FUNCTION_BLOCK FB_ProcessControl

VAR_IN_OUT
	stProcessControl	:	ST_ProcessControl	;
END_VAR
VAR
	bRun			: BOOL	;
	//fbPID	: 	FB_BasicPID	;
	fbPID	: 	PID	;
	hystCIP_SetPoint: FB_Hysteresis_REAL;
	Call_ActDelayTON	: TON	;
	bRunCalled		: BOOL	;//mRun was called since the last body call

	handling_PID_Manual: TON;

END_VAR

//stProcessControl.bManual:=TRUE;



//Deactivate control 1s after mRun stops being called (body may be called several times per cycle)
Call_ActDelayTON(IN:=stProcessControl.bActiveCntr AND NOT bRunCalled , PT:=T#1S , Q=> , ET=> );
bRunCalled:=FALSE;

m_Check();

act_Call_PID();
act_CallHyst();

handling_PID_Manual(PT:=T#0.5S);//, IN:=TRUE
IF handling_PID_Manual.Q THEN;
	stProcessControl.bManual:=TRUE;
ELSE;
	stProcessControl.bManual:=FALSE;
END_IF

ACTION act_Call_PID:
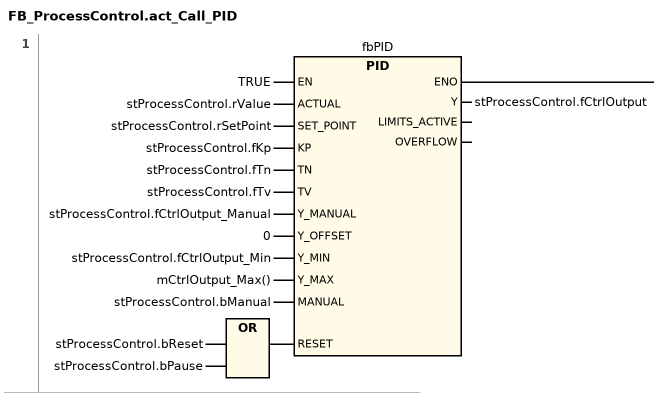
// NETWORK 1
fbPID(
    ACTUAL := stProcessControl.rValue,
    SET_POINT := stProcessControl.rSetPoint,
    KP := stProcessControl.fKp,
    TN := stProcessControl.fTn,
    TV := stProcessControl.fTv,
    Y_MANUAL := stProcessControl.fCtrlOutput_Manual,
    Y_OFFSET := 0,
    Y_MIN := stProcessControl.fCtrlOutput_Min,
    Y_MAX := mCtrlOutput_Max(),
    MANUAL := stProcessControl.bManual,
    RESET := stProcessControl.bReset OR stProcessControl.bPause,
    Y => stProcessControl.fCtrlOutput); // PID
END_ACTION

ACTION act_Call_PID_old:

	
(*
fbPID(
	fSetpointValue:=stProcessControl.rSetPoint , 
	fActualValue:=stProcessControl.rValue , 
	bReset:=stProcessControl.bReset , 
	fCtrlCycleTime:=stProcessControl.fCtrlCycleTime , 
	fKp:=stProcessControl.fKp , 
	fTn:=stProcessControl.fTn , 
	fTv:=stProcessControl.fTv , 
	fTd:=stProcessControl.fTd , 
	fCtrlOutput=>stProcessControl.fCtrlOutput , 
	nErrorStatus=>stProcessControl.nErrorStatus );
*)
END_ACTION

ACTION act_CallHyst:
hystCIP_SetPoint(
	fIn:=stProcessControl.rValue,//g_HMI.stT4_Sens.rTankLevel,
	fHigh:=stProcessControl.fHystHigh,
	fLow:=stProcessControl.fHystLow,
	iDigitsAfterDot:=,
	bOut=>stProcessControl.bHystOut);
END_ACTION

METHOD m_Check : BOOL
VAR_INPUT
END_VAR
IF NOT __ISVALIDREF(stProcessControl) THEN
	RETURN;
END_IF

IF bRun THEN
	stProcessControl.bActiveCntr:=TRUE;
	bRunCalled:=TRUE;
ELSIF NOT bRun AND Call_ActDelayTON.Q THEN
	stProcessControl.bActiveCntr:=FALSE;
END_IF

IF bRun THEN
	stProcessControl.Deviation:=stProcessControl.rSetPoint-stProcessControl.rValue;
	stProcessControl.Control_ON:=FALSE;
	stProcessControl.OverFlow:=FALSE;
	stProcessControl.bDone:=FALSE;
	
	IF stProcessControl.Deviation >= stProcessControl.ToleravceLow THEN;
		//Value too low needs to be increased
		stProcessControl.Control_ON:=TRUE;
		stProcessControl.OverFlow:=FALSE;
		stProcessControl.bDone:=FALSE;
	ELSIF stProcessControl.Deviation <= -stProcessControl.ToleranceHigh THEN;
		//value too high need to be decreased
		stProcessControl.OverFlow:=TRUE;
		stProcessControl.Control_ON:=TRUE;
		stProcessControl.bDone:=FALSE;
		//message
	ELSE;
		// Done, value in tolerace
		stProcessControl.OverFlow:=FALSE;
		stProcessControl.Control_ON:=FALSE;
		stProcessControl.bDone:=TRUE;
	END_IF
	bRun:=FALSE;
END_IF
END_METHOD

METHOD mCtrlOutput_Max : REAL
VAR_INPUT
END_VAR

VAR
	span: LREAL;
END_VAR


span:=ABS(stProcessControl.fCtrlOutput_Max-stProcessControl.fCtrlOutput_Min);
//LimitedPrecentage:=
IF stProcessControl.rValue>stProcessControl.rValue_Min_To_ReleaseControl THEN;
	mCtrlOutput_Max:=stProcessControl.fCtrlOutput_Max;
ELSE;
	mCtrlOutput_Max:=stProcessControl.fCtrlOutput_Min+(span*0.3);
END_IF
END_METHOD

METHOD mManual : BOOL
VAR_INPUT
	value: BOOL;
END_VAR
//PID manual request without starting control (bRun/bActiveCntr untouched)
handling_PID_Manual(IN:=value);
mManual:=stProcessControl.bManual;
END_METHOD

METHOD mPause : BOOL
VAR_INPUT
	value: BOOL;
END_VAR
stProcessControl.bPause:=value;
END_METHOD

METHOD mReset : BOOL
VAR_INPUT
END_VAR
stProcessControl.Control_ON:=FALSE;
stProcessControl.OverFlow:=FALSE;
stProcessControl.bDone:=FALSE;
END_METHOD

METHOD mRun : BOOL
VAR_INPUT
	//Set_Point: REAL;
END_VAR
bRun:=TRUE;
//stProcessControl.rSetPoint:=Set_Point;
m_Check();



mRun:=stProcessControl.bDone;
END_METHOD

METHOD mRun_Hyst : REAL
VAR_INPUT
END_VAR
stProcessControl.bManual:=FALSE;
IF stProcessControl.bHystOut THEN
	mRun_Hyst:=stProcessControl.rHystOutLow;
ELSE
	mRun_Hyst:=stProcessControl.rHystOutHigh;
END_IF
END_METHOD

METHOD mRun_PID : REAL
VAR_INPUT
	Set_Point: REAL;
	controlManual: BOOL;
END_VAR
mRun();//mRun(Set_Point:=Set_Point);
//stProcessControl.bManual:=controlManual;
//stProcessControl.rSetPoint:=Set_Point;
handling_PID_Manual(IN:=controlManual);
mRun_PID:=stProcessControl.fCtrlOutput;
END_METHOD

METHOD mRun_With_SP : BOOL
VAR_INPUT
	Set_Point: REAL;
END_VAR
stProcessControl.rSetPoint:=Set_Point;
bRun:=TRUE;
mRun();
//stProcessControl.rSetPoint:=Set_Point;
mRun_With_SP:=stProcessControl.bDone;
END_METHOD

END_FUNCTION_BLOCK

(* stored: Version 1.1.0.1, ProductVersion 3.1.4026.21
   POU FB_ProcessControl: Id {a1972051-d534-4d79-bd7a-71cd1b516897}, SpecialFunc None
   Action act_Call_PID: Id {839fbd4c-e468-439d-b2e8-fa15b4ee659a}
   Action act_Call_PID_old: Id {e29ea305-112b-4479-9e5c-3d503fcea5b6}
   Action act_CallHyst: Id {7f4572c7-9e9a-4bff-b0e0-f6c19cca19c6}
   Method m_Check: Id {b27ec81e-04ce-483d-958b-1ee4b2519c56}
   Method mCtrlOutput_Max: Id {96e0187b-897b-496a-b800-2f20b878b88c}
   Method mManual: Id {1beeeb9a-e732-4638-8ad0-65b51ae96f3a}
   Method mPause: Id {be53090d-a73d-45ab-9fd1-26dc14e563ed}
   Method mReset: Id {b49576d6-978e-47f7-ae59-752a1612df43}
   Method mRun: Id {9603e267-93ce-4898-8d8d-2a4ace5f7fdf}
   Method mRun_Hyst: Id {ddfa5b4a-f749-4a9f-b8a9-9760265fd642}
   Method mRun_PID: Id {4a3f5dec-9850-4133-86e5-b2ae6f3c1d56}
   Method mRun_With_SP: Id {2d03209f-e46c-40c1-b393-0560a9377f6a} *)
